FUNCTION_BLOCK FB_ToggleBit
VAR_INPUT
(*+++++ TxPDO Toggle +++++*)
	bToggle: BOOL;
END_VAR
VAR_OUTPUT
END_VAR
VAR
(*+++++ Toggle Bit Bridge +++++*)
	rtToggle: R_TRIG;
	ftToggle: F_TRIG;
	rCounter: REAL;
	rLastCounter: REAL;
(*+++++ Evaluation of Toggle Bits +++++*)
	tonTimer: TON;
	rToggleBitCounter: REAL;
	rUpdateTime: REAL;
END_VAR

(*This function block evaluates the Toggle Bit of the device.
Within a period of 10 seconds, is is checked how often the Toggle Bit changes it's value. *)

rtToggle(CLK:= bToggle);
ftToggle(CLK:= bToggle);

tonTimer.IN:= TRUE;
tonTimer.PT:= t#10000ms;

IF NOT tonTimer.Q THEN
	IF rtToggle.Q THEN
		rCounter:= rCounter+1;
	END_IF
	IF ftToggle.Q THEN
		rCounter:= rCounter+1;
	END_IF

	rToggleBitCounter:= rCounter;
ELSE
	rLastCounter:= rCounter;
	rUpdateTime:= 1/ (rLastCounter/10); 		(*Update Time is calculated*)
	rCounter:= 0;
	tonTimer.IN:= FALSE;
END_IF

tonTimer();

END_FUNCTION_BLOCK

(* stored: Version 1.1.0.1, ProductVersion 3.1.4024.15
   POU FB_ToggleBit: Id {397c6029-8a54-4af3-9835-5d1d28359bb5}, SpecialFunc None *)
